(* IEC 61131-3 sources: RVM_Dijital_Ikiz_ModelveOtomasyon_BitirmeProjesi/Codesys_Dosyalari/Paylasim/PLC_Kaynaklari, 10 files *)

(* ---- FB_CikisKontrolLD_decl.st ---- *)
FUNCTION_BLOCK FB_CikisKontrolLD
VAR_INPUT
    // Diagnostic inputs: confirm scan updates without changing ladder logic.
    udiCevrimNo : UDINT;
    uiMakineDurumu : UINT;
	xCalismaIzni: BOOL;
	xBaglanti: BOOL;
	xVeriGecerli: BOOL;
	xAcilStop: BOOL;
	xSikisma: BOOL;
	xDurdur: BOOL;
	xGirisAsamasi: BOOL;
	xKabulAsamasi: BOOL;
	xIadeAsamasi: BOOL;
	xKirmaAsamasi: BOOL;
	xHazneAsamasi: BOOL;
	xEveDonusAsamasi: BOOL;
	xBosaltmaAsamasi: BOOL;
	xTanimaOnayi: BOOL;
	xKapakKapali: BOOL;
	xHedefte: BOOL;
END_VAR
VAR_OUTPUT
	xHareketIzni: BOOL;
	xIleriIstegi: BOOL;
	xGeriIstegi: BOOL;
	xKiriciCalis: BOOL;
	xHazneHareket: BOOL;
	xKapakAc: BOOL;
END_VAR

(* ---- FB_KomutOnceligi106_decl.st ---- *)
FUNCTION_BLOCK FB_KomutOnceligi106
VAR_INPUT
    uiKomutKodu : UINT;
    xYeniKomut : BOOL;
    udiKomutKimligi : UDINT;
END_VAR
VAR_OUTPUT
    uiOncelik : UINT;
    udiCevrimSayaci : UDINT;
    uiSonKomutKodu : UINT;
    uiSonOncelik : UINT;
    udiSonKomutKimligi : UDINT;
END_VAR

(* ---- FB_KonveyorIzin_decl.st ---- *)
FUNCTION_BLOCK FB_KonveyorIzin
VAR_INPUT
    xIzin        : BOOL;
    xIleriIstegi : BOOL;
    xGeriIstegi  : BOOL;
END_VAR
VAR_OUTPUT
    xIleri        : BOOL;
    xGeri         : BOOL;
    xYonCakismasi : BOOL;
END_VAR

(* ---- FB_MalzemeSiniflandirma106_decl.st ---- *)
FUNCTION_BLOCK FB_MalzemeSiniflandirma106
VAR_INPUT
    rMetal : REAL;
    rManyetik : REAL;
    rKutleGram : REAL;
    rGecirgenlik : REAL;
    rYansima : REAL;
    rBoyMetre : REAL;
    rEnMetre : REAL;
    rDoluluk : REAL;
    xVeriYasiUygun : BOOL := TRUE;
    xSensorlerGecerli : BOOL := TRUE;
    xSekilUygun : BOOL := TRUE;
    udiUrunKimligi : UDINT;
    udiPlcOturumu : UDINT;
    udiUnityOturumu : UDINT;
    udiGoruntuIstegi : UDINT;
END_VAR
VAR_OUTPUT
    xDegerlendirildi : BOOL;
    udiDegerlendirmeSayaci : UDINT;
    uiMalzeme : UINT;
    uiGoruntuKarari : UINT;
    uiRetNedeni : UINT;
    rBoyCm : REAL;
    rEnCm : REAL;
    rYuzeyAlani : REAL;
    rHacim : REAL;
    rKabukYogunluk : REAL;
    rHacimYogunluk : REAL;
    xTemelSinirlarUygun : BOOL;
    xAlanUygun : BOOL;
    xPetKosullari : BOOL;
    xCamKosullari : BOOL;
    xAluminyumKosullari : BOOL;
    xMetalBelirsiz : BOOL;
END_VAR

(* ---- FB_RVMControl106_decl.st ---- *)
FUNCTION_BLOCK FB_RVMControl106
VAR_INPUT
    inp : ST_RVMInput106;
    op : ST_RVMOperator106;
    fresh : BOOL;
    epoch : UDINT;
END_VAR
VAR_OUTPUT
    q : ST_RVMOutput106;
END_VAR
VAR
    a : ST_RVMInput106;
    initialized : BOOL;
    session : UDINT;
    packet : UDINT;
    heartbeat : BOOL;
    synchronized : BOOL;
    sessionChanged : BOOL;
    dataOK : BOOL;
    linked : BOOL;
    home : BOOL;
    emptyHome : BOOL;
    emergency : BOOL;
    stopLevel : BOOL;
    targetFull : BOOL;
    faultNow : UINT;
    previousState : UINT;
    previousButtons : ARRAY[1..5] OF BOOL;
    armed : ARRAY[1..5] OF BOOL;
    buttons : ARRAY[1..5] OF BOOL;
    edges : ARRAY[1..5] OF BOOL;
    newRequest : ARRAY[1..2] OF BOOL;
    cmdId : ARRAY[1..2] OF UDINT;
    cmdCode : ARRAY[1..2] OF UINT;
    cmdParam : ARRAY[1..2] OF UINT;
    cachedStatus : ARRAY[1..2] OF UINT;
    cachedReason : ARRAY[1..2] OF UINT;
    replyId : ARRAY[1..2] OF UDINT;
    replyStatus : ARRAY[1..2] OF UINT;
    replyReason : ARRAY[1..2] OF UINT;
    source : INT;
    chosen : INT;
    other : INT;
    i : INT;
    hmiCode : UINT;
    hmiParam : UINT;
    resultStatus : UINT;
    resultReason : UINT;
    pendingSource : INT;
    pendingId : UDINT;
    insertConfirmed : BOOL;
    confirmedProduct : UDINT;
    lastProduct : UDINT;
    waitLink : TON;
    waitStage : TON;
    waitRecognition : TON;
    waitVision : TON;
    visionMatch : BOOL;
    visionShape : BOOL;
    waitCycle : TON;
    waitInsert : TON;
    fbMalzeme : FB_MalzemeSiniflandirma106;
    fbUnityOncelik : FB_KomutOnceligi106;
    fbCodesysOncelik : FB_KomutOnceligi106;
    fbCikisLD : FB_CikisKontrolLD;
    fbKonveyorIzin : FB_KonveyorIzin;
END_VAR

(* ---- FB_KomutOnceligi106_body.st ---- *)
// Same command priorities; separate instances for Unity and CODESYS HMI.
CASE uiKomutKodu OF
2: uiOncelik := 1;
3: uiOncelik := 2;
5: uiOncelik := 3;
1: uiOncelik := 4;
4: uiOncelik := 5;
ELSE uiOncelik := 99;
END_CASE;
IF udiCevrimSayaci = UDINT#4294967295 THEN
    udiCevrimSayaci := 1;
ELSE
    udiCevrimSayaci := udiCevrimSayaci + 1;
END_IF;
IF xYeniKomut THEN
    uiSonKomutKodu := uiKomutKodu;
    uiSonOncelik := uiOncelik;
    udiSonKomutKimligi := udiKomutKimligi;
END_IF;

(* ---- FB_MalzemeSiniflandirma106_body.st ---- *)
// Last completed classification attempt. Inputs and results remain visible.
// Each attempt clears intermediate values, including early rejection paths.
xDegerlendirildi := TRUE;
IF udiDegerlendirmeSayaci = UDINT#4294967295 THEN
    udiDegerlendirmeSayaci := 1;
ELSE
    udiDegerlendirmeSayaci := udiDegerlendirmeSayaci + 1;
END_IF;
uiMalzeme := 0; uiGoruntuKarari := 2; uiRetNedeni := 0;
rBoyCm := 0; rEnCm := 0; rYuzeyAlani := 0; rHacim := 0;
rKabukYogunluk := 0; rHacimYogunluk := 0;
xTemelSinirlarUygun := FALSE; xAlanUygun := FALSE;
xPetKosullari := FALSE; xCamKosullari := FALSE;
xAluminyumKosullari := FALSE; xMetalBelirsiz := FALSE;

// Same order as the previous controller guards.
IF NOT xVeriYasiUygun THEN uiRetNedeni := 10; uiGoruntuKarari := 4; RETURN; END_IF;
IF NOT xSensorlerGecerli THEN uiRetNedeni := 11; uiGoruntuKarari := 3; RETURN; END_IF;
IF NOT xSekilUygun THEN uiRetNedeni := 12; RETURN; END_IF;

xTemelSinirlarUygun := (rMetal>=0) AND (rMetal<=1) AND (rManyetik>=0) AND (rManyetik<=0.1)
    AND (rKutleGram>=5) AND (rKutleGram<=1000) AND (rGecirgenlik>=0) AND (rGecirgenlik<=1)
    AND (rYansima>=0) AND (rYansima<=1) AND (rBoyMetre>=0.10) AND (rBoyMetre<=0.30)
    AND (rEnMetre>=0.02) AND (rEnMetre<=0.09) AND (rDoluluk>0) AND (rDoluluk<=1);
IF NOT xTemelSinirlarUygun THEN uiRetNedeni := 1; RETURN; END_IF;
rBoyCm := rBoyMetre * 100.0;
rEnCm := rEnMetre * 100.0;
rYuzeyAlani := 3.14159265 * rEnCm * rBoyCm * rDoluluk;
xAlanUygun := rYuzeyAlani > 1.0;
IF NOT xAlanUygun THEN uiRetNedeni := 2; RETURN; END_IF;
rHacim := rYuzeyAlani * rEnCm / 4.0;
rKabukYogunluk := rKutleGram / rYuzeyAlani;
rHacimYogunluk := rKutleGram / rHacim;

xAluminyumKosullari := (rMetal>=0.5) AND (rGecirgenlik<=0.08)
    AND (rKutleGram>=8) AND (rKutleGram<=45) AND (rBoyMetre<=0.20);
xPetKosullari := (rMetal<=0.1) AND (rKutleGram>=8) AND (rKutleGram<=75)
    AND (rKabukYogunluk>=0.040) AND (rKabukYogunluk<=0.095) AND (rGecirgenlik>=0.35);
xCamKosullari := (rMetal<=0.1) AND (rKutleGram>=100) AND (rKutleGram<=800)
    AND (rKabukYogunluk>=0.450) AND (rKabukYogunluk<=0.680) AND (rDoluluk>=0.875)
    AND (rGecirgenlik>=0.45) AND (rGecirgenlik<=0.85) AND (rYansima>=0.12);
xMetalBelirsiz := (rMetal>0.1) AND (rMetal<0.5);
IF rMetal>=0.5 THEN
    IF xAluminyumKosullari THEN uiMalzeme := 2; ELSE uiRetNedeni := 3; END_IF;
ELSIF rMetal<=0.1 THEN
    IF xPetKosullari THEN uiMalzeme := 1;
    ELSIF xCamKosullari THEN uiMalzeme := 3;
    ELSE uiRetNedeni := 5;
    END_IF;
ELSE
    uiRetNedeni := 4;
END_IF;
IF uiMalzeme<>0 THEN uiGoruntuKarari := 1; END_IF;

(* ---- FB_RVMControl106_body.st ---- *)
// Single process owner. No actuator command is derived from a UI bit directly.
q.uiProtokolSurumu := 106;
q.udiPlcOturumu := epoch;
q.uiDesteklenenModlar := 2; // Render camera + simulated physical sensors only.
q.uiVeriModu := 1;
q.rBantHizi := 0.85;
q.rKiriciDevri := 120.0;
q.rHazneHizi := 1.5;
q.rKapakAcisi := 75.0;
q.udiPlcSayaci := q.udiPlcSayaci + 1;
heartbeat := FALSE;
sessionChanged := FALSE;
newRequest[1] := FALSE;
newRequest[2] := FALSE;
insertConfirmed := FALSE;
faultNow := 0;
IF NOT initialized THEN
    initialized := TRUE;
    q.uiDurum := 0;
    q.xCalismaIzni := FALSE;
    q.rHazneHedefi := 0.225;
END_IF;
IF epoch = 0 THEN faultNow := 313; END_IF;

// A zero-epoch HELLO is mandatory before this PLC incarnation accepts commands.
// The HELLO'inp command watermark is consumed, never executed.
IF fresh AND (inp.udiUnityOturumu <> 0) AND (inp.udiUnitySayaci <> 0) THEN
    IF (inp.udiGorulenPlcOturumu = 0) AND ((session <> inp.udiUnityOturumu) OR NOT synchronized) THEN
        a := inp;
        sessionChanged := session <> inp.udiUnityOturumu;
        session := inp.udiUnityOturumu;
        lastProduct := 0;
        packet := inp.udiUnitySayaci;
        synchronized := TRUE;
        cmdId[1] := inp.udiKomutKimligi;
        cmdCode[1] := inp.uiOperatorKomutu;
        cmdParam[1] := inp.uiOperatorParametresi;
        cachedStatus[1] := 5;
        cachedReason[1] := 10;
        replyId[1] := cmdId[1];
        replyStatus[1] := 5;
        replyReason[1] := 10;
        q.xCalismaIzni := FALSE;
        IF q.uiHataKodu = 0 THEN q.uiDurum := 0; END_IF;
    ELSIF synchronized AND (session = inp.udiUnityOturumu)
        AND (inp.udiGorulenPlcOturumu = epoch) AND (inp.udiUnitySayaci > packet) THEN
        packet := inp.udiUnitySayaci;
        a := inp;
        heartbeat := TRUE;
        IF inp.udiKomutKimligi > cmdId[1] THEN
            cmdId[1] := inp.udiKomutKimligi;
            cmdCode[1] := inp.uiOperatorKomutu;
            cmdParam[1] := inp.uiOperatorParametresi;
            newRequest[1] := TRUE;
        ELSIF (inp.udiKomutKimligi <> cmdId[1]) OR (inp.uiOperatorKomutu <> cmdCode[1])
            OR (inp.uiOperatorParametresi <> cmdParam[1]) THEN
            replyId[1] := inp.udiKomutKimligi;
            replyStatus[1] := 3;
            replyReason[1] := 13;
        ELSE
            replyId[1] := cmdId[1];
            replyStatus[1] := cachedStatus[1];
            replyReason[1] := cachedReason[1];
        END_IF;
    END_IF;
END_IF;
q.udiUnityOnayOturumu := session;
waitLink(IN := NOT heartbeat, PT := T#750MS);
linked := synchronized AND (session = a.udiUnityOturumu) AND (a.udiGorulenPlcOturumu = epoch)
    AND (epoch <> 0) AND NOT waitLink.Q AND (a.uiUnityProtokol = 106);
home := ABS(a.rHazneKonumu - 0.225) < 0.008;
emptyHome := a.xYolBos AND NOT a.xGiris AND a.xKapakKapali AND NOT a.xKapakAcik AND home;
emergency := op.xAcilStop OR a.xAcilStop;
// Comparisons reject NaN as well as out-of-range values. No invalid data fallback.
dataOK := a.xPlantVerisiGecerli AND (a.uiPlantVeriKaynagi = 1)
    AND (a.rHazneKonumu >= -0.770001) AND (a.rHazneKonumu <= 0.310001)
    AND (a.rKutleGram >= 0.0) AND (a.rKutleGram <= 10000.0)
    AND (a.rBoyMetre >= 0.0) AND (a.rBoyMetre <= 2.000001)
    AND (a.rOptikGecirgenlik >= 0.0) AND (a.rOptikGecirgenlik <= 1.000001)
    AND (a.rGercekBantHizi >= -1.200001) AND (a.rGercekBantHizi <= 1.200001)
    AND (a.rGercekKiriciDevri >= 0.0) AND (a.rGercekKiriciDevri <= 180.0001)
    AND NOT (a.xKapakAcik AND a.xKapakKapali)
    AND NOT (a.xYolBos AND a.xGiris) AND (a.uiBosaltilanKutu <= 3);

// HMI: arm only after FALSE has been observed; held or startup TRUE cannot repeat.
buttons[1] := op.xBaslat; buttons[2] := op.xDurdur; buttons[3] := op.xSifirla;
buttons[4] := op.xNesneEkle; buttons[5] := op.xModUygula;
FOR i := 1 TO 5 DO
    IF NOT buttons[i] THEN armed[i] := TRUE; END_IF;
    edges[i] := armed[i] AND buttons[i] AND NOT previousButtons[i];
    previousButtons[i] := buttons[i];
END_FOR;
hmiCode := 0; hmiParam := 0;
IF edges[2] THEN hmiCode := 2;
ELSIF edges[3] THEN hmiCode := 3;
ELSIF edges[5] THEN hmiCode := 5; hmiParam := op.uiSeciliMod;
ELSIF edges[1] THEN hmiCode := 1;
ELSIF edges[4] THEN hmiCode := 4; hmiParam := op.uiSeciliNesne;
END_IF;
IF hmiCode <> 0 THEN
    IF cmdId[2] = UDINT#4294967295 THEN faultNow := 313;
    ELSE
        cmdId[2] := cmdId[2] + 1;
        cmdCode[2] := hmiCode; cmdParam[2] := hmiParam;
        newRequest[2] := TRUE;
    END_IF;
END_IF;
stopLevel := op.xDurdur OR (newRequest[1] AND (cmdCode[1] = 2));

// Fault priority is stable; reconnecting Unity never clears a latched fault.
IF q.xCalismaIzni THEN
    IF emergency THEN faultNow := 303;
    // Unity also raises its local motion interlock on an identity mismatch.
    // Preserve the specific cause while the session is valid, before generic jam/data flags.
    ELSIF linked AND (q.uiDurum >= 20) AND (q.uiDurum <= 100) AND (a.udiUrunKimligi <> q.udiIslemKimligi) THEN faultNow := 305;
    ELSIF a.xSikisma THEN faultNow := 304;
    ELSIF a.uiUnityProtokol <> 106 THEN faultNow := 302;
    ELSIF NOT linked THEN faultNow := 301;
    ELSIF NOT dataOK THEN faultNow := 310;
    END_IF;
END_IF;
waitStage(IN := (q.uiDurum = previousState) AND (q.uiDurum >= 20) AND (q.uiDurum <= 100), PT := T#8S);
previousState := q.uiDurum;
waitRecognition(IN := q.uiDurum = 30, PT := T#200MS);
waitVision(IN := q.uiDurum = 30, PT := T#4S);
visionMatch := (a.udiGoruntuOnayi = q.udiGoruntuIstegi) AND (q.udiGoruntuIstegi <> 0)
    AND (a.udiGoruntuUrunu = q.udiIslemKimligi) AND (a.udiGoruntuPlcOturumu = epoch)
    AND (a.udiGoruntuUnityOturumu = session);
visionShape := a.xGoruntuNesneVar AND (a.rGoruntuBoy >= 0.10) AND (a.rGoruntuBoy <= 0.30)
    AND (a.rGoruntuEn >= 0.02) AND (a.rGoruntuEn <= 0.09)
    AND (a.rGoruntuBoy >= 1.5*a.rGoruntuEn) AND (a.rGoruntuBoy <= 7.0*a.rGoruntuEn)
    AND (a.rGoruntuDoluluk >= 0.35) AND (a.rGoruntuDoluluk <= 1.0);
waitCycle(IN := (q.uiDurum >= 20) AND (q.uiDurum <= 90), PT := T#5600MS);
waitInsert(IN := q.xNesneIstegiEtkin, PT := T#2S);
IF waitStage.Q AND (faultNow = 0) THEN faultNow := 306; END_IF;
IF faultNow <> 0 AND q.uiHataKodu = 0 THEN q.uiHataKodu := faultNow; END_IF;
IF stopLevel OR emergency OR sessionChanged OR (q.uiHataKodu <> 0) THEN
    q.xCalismaIzni := FALSE;
    IF q.uiHataKodu = 0 THEN q.uiDurum := 0; ELSE q.uiDurum := 900; END_IF;
    IF q.xNesneIstegiEtkin THEN
        cachedStatus[pendingSource] := 5; cachedReason[pendingSource] := 1;
        IF replyId[pendingSource] = pendingId THEN
            replyStatus[pendingSource] := 5; replyReason[pendingSource] := 1;
        END_IF;
    END_IF;
    q.xNesneIstegiEtkin := FALSE;
END_IF;

// Arbitration is deterministic. No deferred queue can start work after a stop.
fbUnityOncelik(uiKomutKodu := cmdCode[1], xYeniKomut := newRequest[1], udiKomutKimligi := cmdId[1]);
fbCodesysOncelik(uiKomutKodu := cmdCode[2], xYeniKomut := newRequest[2], udiKomutKimligi := cmdId[2]);
chosen := 0;
IF newRequest[2] THEN chosen := 2; END_IF;
IF newRequest[1] THEN
    IF chosen = 0 THEN chosen := 1;
    ELSIF fbUnityOncelik.uiOncelik < fbCodesysOncelik.uiOncelik THEN chosen := 1;
    END_IF;
END_IF;
FOR source := 1 TO 2 DO
    IF newRequest[source] THEN
        resultStatus := 3; resultReason := 0;
        replyId[source] := cmdId[source];
        IF (source <> chosen) AND NOT (cmdCode[source] = 2) THEN
            IF stopLevel THEN resultReason := 1; ELSE resultReason := 9; END_IF;
        ELSIF cmdCode[source] = 2 THEN
            q.xCalismaIzni := FALSE;
            IF q.uiHataKodu = 0 THEN q.uiDurum := 0; ELSE q.uiDurum := 900; END_IF;
            resultStatus := 2;
        ELSIF (cmdCode[source] = 0) OR (cmdCode[source] > 5)
            OR ((cmdCode[source] <= 3) AND (cmdParam[source] <> 0))
            OR ((cmdCode[source] = 4) AND (cmdParam[source] > 3))
            OR ((cmdCode[source] = 5) AND (cmdParam[source] > 2)) THEN resultReason := 7;
        ELSIF stopLevel THEN resultReason := 1;
        ELSIF emergency OR a.xSikisma THEN resultReason := 5;
        ELSIF NOT linked OR NOT dataOK THEN resultReason := 2;
        ELSIF q.xNesneIstegiEtkin THEN resultReason := 6;
        ELSE
            CASE cmdCode[source] OF
            1:
                IF q.uiHataKodu <> 0 THEN resultReason := 5;
                ELSIF q.uiDurum <> 0 THEN resultReason := 3;
                ELSIF NOT emptyHome THEN resultReason := 4;
                ELSE q.xCalismaIzni := TRUE; q.uiDurum := 10; resultStatus := 2;
                END_IF;
            3:
                IF q.xCalismaIzni OR ((q.uiDurum <> 0) AND (q.uiDurum <> 900)) THEN resultReason := 3;
                ELSIF NOT emptyHome THEN resultReason := 4;
                ELSIF epoch = 0 THEN resultReason := 10;
                ELSE q.uiHataKodu := 0; q.uiDurum := 0; q.xCalismaIzni := FALSE; resultStatus := 2;
                END_IF;
            4:
                IF q.uiHataKodu <> 0 THEN resultReason := 5;
                ELSIF (q.uiDurum <> 10) OR NOT q.xCalismaIzni THEN resultReason := 3;
                ELSIF NOT emptyHome THEN resultReason := 4;
                ELSIF q.udiNesneIstegi = UDINT#4294967295 THEN resultReason := 10;
                ELSE
                    q.udiNesneIstegi := q.udiNesneIstegi + 1;
                    q.uiNesneProfili := cmdParam[source];
                    q.xNesneIstegiEtkin := TRUE;
                    pendingSource := source; pendingId := cmdId[source];
                    resultStatus := 1;
                END_IF;
            5:
                IF cmdParam[source] <> 1 THEN resultReason := 8;
                ELSIF (q.uiDurum <> 0) OR q.xCalismaIzni THEN resultReason := 3;
                ELSIF NOT emptyHome THEN resultReason := 4;
                ELSE q.uiVeriModu := 1; resultStatus := 2;
                END_IF;
            END_CASE;
        END_IF;
        cachedStatus[source] := resultStatus; cachedReason[source] := resultReason;
        replyStatus[source] := resultStatus; replyReason[source] := resultReason;
        IF source = chosen THEN q.uiSonKomutKaynagi := INT_TO_UINT(source); END_IF;
    END_IF;
END_FOR;

// Product admission is tied to the PLC-issued request, not just a presence bit.
IF q.xNesneIstegiEtkin THEN
    resultStatus := 1; resultReason := 0;
    IF waitInsert.Q THEN
        resultStatus := 4; resultReason := 11;
        q.uiHataKodu := 312; // A delayed physical creation must require explicit recovery.
    ELSIF heartbeat AND (a.udiNesneOnayi = q.udiNesneIstegi) THEN
        IF a.uiNesneSonucu = 2 THEN resultStatus := 3; resultReason := 12;
        ELSIF a.uiNesneSonucu = 1 THEN
            IF (a.udiNesneUrunKimligi <> 0) AND (a.udiNesneUrunKimligi = a.udiUrunKimligi)
                AND (a.udiUrunKimligi > lastProduct) AND a.xGiris AND NOT a.xYolBos THEN
                confirmedProduct := a.udiUrunKimligi;
                lastProduct := a.udiUrunKimligi;
                insertConfirmed := TRUE;
                resultStatus := 2;
            ELSE resultStatus := 3; resultReason := 12; q.uiHataKodu := 312;
            END_IF;
        END_IF;
    END_IF;
    IF resultStatus <> 1 THEN
        q.xNesneIstegiEtkin := FALSE;
        IF cmdId[pendingSource] = pendingId THEN
            cachedStatus[pendingSource] := resultStatus; cachedReason[pendingSource] := resultReason;
        END_IF;
        IF replyId[pendingSource] = pendingId THEN
            replyStatus[pendingSource] := resultStatus; replyReason[pendingSource] := resultReason;
        END_IF;
    END_IF;
END_IF;

targetFull := ((q.uiHedefKutu = 1) AND a.xKutuPetDolu)
    OR ((q.uiHedefKutu = 2) AND a.xKutuAluminyumDolu)
    OR ((q.uiHedefKutu = 3) AND a.xKutuCamDolu);
IF q.xCalismaIzni AND (q.uiDurum >= 40) AND (q.uiDurum <= 70) AND targetFull THEN q.uiHataKodu := 308; END_IF;
IF q.uiHataKodu = 0 AND q.xCalismaIzni THEN
    CASE q.uiDurum OF
    10:
        q.xTanimaOnayi := FALSE; q.uiTaninmisMalzeme := 0; q.uiHedefKutu := 0;
        IF insertConfirmed THEN q.udiIslemKimligi := confirmedProduct; q.uiDurum := 20;
        ELSIF NOT a.xYolBos AND NOT q.xNesneIstegiEtkin THEN q.uiHataKodu := 312;
        END_IF;
    20:
        IF a.xTanima THEN
            IF q.udiGoruntuIstegi = UDINT#4294967295 THEN q.uiHataKodu := 313;
            ELSE q.udiGoruntuIstegi := q.udiGoruntuIstegi+1; q.uiGoruntuKarari := 0; q.uiDurum := 30;
            END_IF;
        END_IF;
    30:
        IF NOT a.xTanima THEN q.uiHataKodu := 307;
        ELSIF waitVision.Q THEN
            q.uiGoruntuKarari := 5; q.uiTaninmisMalzeme := 0; q.uiHedefKutu := 0; q.uiDurum := 100;
        ELSIF waitRecognition.Q AND visionMatch THEN
            q.uiTaninmisMalzeme := 0;
            fbMalzeme(
                rMetal := a.rOlcumMetal, rManyetik := a.rOlcumManyetik,
                rKutleGram := a.rKutleGram, rGecirgenlik := a.rOptikGecirgenlik,
                rYansima := a.rOlcumYansima, rBoyMetre := a.rGoruntuBoy,
                rEnMetre := a.rGoruntuEn, rDoluluk := a.rGoruntuDoluluk,
                xVeriYasiUygun := (a.rGoruntuYasiMs >= 0.0) AND (a.rGoruntuYasiMs <= 2000.0),
                xSensorlerGecerli := a.xGoruntuGecerli AND a.xOlcumTartiGecerli AND a.xOlcumProbGecerli,
                xSekilUygun := visionShape,
                udiUrunKimligi := q.udiIslemKimligi, udiPlcOturumu := epoch,
                udiUnityOturumu := a.udiUnityOturumu, udiGoruntuIstegi := q.udiGoruntuIstegi);
            q.uiTaninmisMalzeme := fbMalzeme.uiMalzeme;
            q.uiGoruntuKarari := fbMalzeme.uiGoruntuKarari;
            q.uiHedefKutu := q.uiTaninmisMalzeme;
            CASE q.uiHedefKutu OF
            1: q.rHazneHedefi := -0.23;
            2: q.rHazneHedefi := -0.77;
            3: q.rHazneHedefi := 0.31;
            END_CASE;
            IF q.uiHedefKutu = 0 THEN q.uiDurum := 100;
            ELSIF ((q.uiHedefKutu=1) AND a.xKutuPetDolu) OR ((q.uiHedefKutu=2) AND a.xKutuAluminyumDolu)
                OR ((q.uiHedefKutu=3) AND a.xKutuCamDolu) THEN q.uiHataKodu := 308;
            ELSE q.xTanimaOnayi := TRUE; q.uiDurum := 40;
            END_IF;
        END_IF;
    40:
        IF NOT a.xKapakKapali THEN q.uiHataKodu := 310;
        ELSIF a.xKiriciGiris THEN q.uiDurum := 50; END_IF;
    50:
        IF a.xKirildi AND a.xHazneDolu AND a.xKapakKapali THEN q.uiDurum := 60; END_IF;
    60:
        IF NOT a.xKapakKapali OR NOT a.xHazneDolu THEN q.uiHataKodu := 310;
        ELSIF ABS(a.rHazneKonumu-q.rHazneHedefi)<0.008 THEN q.uiDurum := 70; END_IF;
    70:
        IF ABS(a.rHazneKonumu-q.rHazneHedefi)>=0.008 THEN q.uiHataKodu := 310;
        ELSIF a.xBosaltildi AND a.xKapakAcik AND NOT a.xHazneDolu AND a.xYolBos THEN
            IF a.uiBosaltilanKutu <> q.uiHedefKutu THEN q.uiHataKodu := 309;
            ELSE q.uiDurum := 80; END_IF;
        END_IF;
    80:
        IF a.xKapakKapali AND NOT a.xKapakAcik AND a.xYolBos AND NOT a.xHazneDolu THEN
            CASE q.uiHedefKutu OF
            1: q.udiPetSayaci := q.udiPetSayaci + 1;
            2: q.udiAluminyumSayaci := q.udiAluminyumSayaci + 1;
            3: q.udiCamSayaci := q.udiCamSayaci + 1;
            END_CASE;
            q.uiDurum := 90;
        END_IF;
    90:
        q.rHazneHedefi := 0.225;
        IF NOT a.xKapakKapali THEN q.uiHataKodu := 310;
        ELSIF home AND a.xYolBos AND waitCycle.Q THEN q.uiDurum := 10; END_IF;
    100:
        IF a.xYolBos THEN q.udiReddedilenSayaci := q.udiReddedilenSayaci+1; q.uiDurum := 10; END_IF;
    END_CASE;
END_IF;

// Apply fault dominance AFTER state processing, in this same scan.
IF q.uiHataKodu <> 0 THEN q.uiDurum := 900; q.xCalismaIzni := FALSE; q.xNesneIstegiEtkin := FALSE; END_IF;
fbCikisLD(
    udiCevrimNo := q.udiPlcSayaci, uiMakineDurumu := q.uiDurum,
    xCalismaIzni := q.xCalismaIzni, xBaglanti := linked, xVeriGecerli := dataOK,
    xAcilStop := emergency, xSikisma := a.xSikisma, xDurdur := stopLevel,
    xGirisAsamasi := q.uiDurum=20, xKabulAsamasi := q.uiDurum=40,
    xIadeAsamasi := q.uiDurum=100, xKirmaAsamasi := q.uiDurum=50,
    xHazneAsamasi := q.uiDurum=60, xEveDonusAsamasi := q.uiDurum=90,
    xBosaltmaAsamasi := q.uiDurum=70, xTanimaOnayi := q.xTanimaOnayi,
    xKapakKapali := a.xKapakKapali, xHedefte := ABS(a.rHazneKonumu-q.rHazneHedefi)<0.008);
fbKonveyorIzin(xIzin := fbCikisLD.xHareketIzni,
    xIleriIstegi := fbCikisLD.xIleriIstegi, xGeriIstegi := fbCikisLD.xGeriIstegi);
q.xKonveyorIleri := fbKonveyorIzin.xIleri;
q.xKonveyorGeri := fbKonveyorIzin.xGeri;
q.xKiriciCalis := fbCikisLD.xKiriciCalis;
q.xHazneHareket := fbCikisLD.xHazneHareket;
q.xKapakAc := fbCikisLD.xKapakAc;
IF NOT q.xCalismaIzni THEN q.xTanimaOnayi := FALSE; END_IF;
q.udiKomutOnayi := replyId[1]; q.uiKomutDurumu := replyStatus[1]; q.uiKomutNedeni := replyReason[1];
q.udiPlcOperatorKomutKimligi := replyId[2]; q.uiPlcOperatorKomutu := cmdCode[2];
q.uiPlcKomutDurumu := replyStatus[2]; q.uiPlcKomutNedeni := replyReason[2];

(* ---- PRG_UnityRVM_body.st ---- *)
IF NOT initialized THEN
    initialized := TRUE;
    IF GVL_RVMKalici.udiOturum < UDINT#4294967295 THEN
        GVL_RVMKalici.udiOturum := GVL_RVMKalici.udiOturum + 1;
        epoch := GVL_RVMKalici.udiOturum;
    END_IF;
END_IF;
fresh := FALSE;
beginMarker := GVL_RVMUnity.udiGirisBaslangic;
IF (beginMarker <> 0) AND (beginMarker = GVL_RVMUnity.udiGirisBitis) AND (beginMarker <> lastMarker) THEN
candidate.uiUnityProtokol := GVL_RVMUnity.uiUnityProtokol;
candidate.udiUnityOturumu := GVL_RVMUnity.udiUnityOturumu;
candidate.udiUnitySayaci := GVL_RVMUnity.udiUnitySayaci;
candidate.udiKomutKimligi := GVL_RVMUnity.udiKomutKimligi;
candidate.uiOperatorKomutu := GVL_RVMUnity.uiOperatorKomutu;
candidate.xGiris := GVL_RVMUnity.xGiris;
candidate.xTanima := GVL_RVMUnity.xTanima;
candidate.xKiriciGiris := GVL_RVMUnity.xKiriciGiris;
candidate.xKirildi := GVL_RVMUnity.xKirildi;
candidate.xHazneDolu := GVL_RVMUnity.xHazneDolu;
candidate.xBosaltildi := GVL_RVMUnity.xBosaltildi;
candidate.xKapakAcik := GVL_RVMUnity.xKapakAcik;
candidate.xKapakKapali := GVL_RVMUnity.xKapakKapali;
candidate.xYolBos := GVL_RVMUnity.xYolBos;
candidate.xMetalAlgilandi := GVL_RVMUnity.xMetalAlgilandi;
candidate.xSikisma := GVL_RVMUnity.xSikisma;
candidate.xAcilStop := GVL_RVMUnity.xAcilStop;
candidate.xKutuPetDolu := GVL_RVMUnity.xKutuPetDolu;
candidate.xKutuAluminyumDolu := GVL_RVMUnity.xKutuAluminyumDolu;
candidate.xKutuCamDolu := GVL_RVMUnity.xKutuCamDolu;
candidate.rKutleGram := GVL_RVMUnity.rKutleGram;
candidate.rOptikGecirgenlik := GVL_RVMUnity.rOptikGecirgenlik;
candidate.rBoyMetre := GVL_RVMUnity.rBoyMetre;
candidate.rHazneKonumu := GVL_RVMUnity.rHazneKonumu;
candidate.rGercekBantHizi := GVL_RVMUnity.rGercekBantHizi;
candidate.rGercekKiriciDevri := GVL_RVMUnity.rGercekKiriciDevri;
candidate.uiBosaltilanKutu := GVL_RVMUnity.uiBosaltilanKutu;
candidate.udiUrunKimligi := GVL_RVMUnity.udiUrunKimligi;
candidate.uiOperatorParametresi := GVL_RVMUnity.uiOperatorParametresi;
candidate.udiGorulenPlcOturumu := GVL_RVMUnity.udiGorulenPlcOturumu;
candidate.udiNesneOnayi := GVL_RVMUnity.udiNesneOnayi;
candidate.uiNesneSonucu := GVL_RVMUnity.uiNesneSonucu;
candidate.udiNesneUrunKimligi := GVL_RVMUnity.udiNesneUrunKimligi;
candidate.uiPlantVeriKaynagi := GVL_RVMUnity.uiPlantVeriKaynagi;
candidate.xPlantVerisiGecerli := GVL_RVMUnity.xPlantVerisiGecerli;
candidate.udiGoruntuOnayi := GVL_RVMUnity.udiGoruntuOnayi;
candidate.udiGoruntuUrunu := GVL_RVMUnity.udiGoruntuUrunu;
candidate.udiGoruntuPlcOturumu := GVL_RVMUnity.udiGoruntuPlcOturumu;
candidate.udiGoruntuUnityOturumu := GVL_RVMUnity.udiGoruntuUnityOturumu;
candidate.xGoruntuGecerli := GVL_RVMUnity.xGoruntuGecerli;
candidate.xGoruntuNesneVar := GVL_RVMUnity.xGoruntuNesneVar;
candidate.rGoruntuBoy := GVL_RVMUnity.rGoruntuBoy;
candidate.rGoruntuEn := GVL_RVMUnity.rGoruntuEn;
candidate.rGoruntuDoluluk := GVL_RVMUnity.rGoruntuDoluluk;
candidate.rGoruntuYasiMs := GVL_RVMUnity.rGoruntuYasiMs;
candidate.xOlcumTartiGecerli := GVL_RVMUnity.xOlcumTartiGecerli;
candidate.xOlcumProbGecerli := GVL_RVMUnity.xOlcumProbGecerli;
candidate.rOlcumYansima := GVL_RVMUnity.rOlcumYansima;
candidate.rOlcumMetal := GVL_RVMUnity.rOlcumMetal;
candidate.rOlcumManyetik := GVL_RVMUnity.rOlcumManyetik;
    fresh := (beginMarker = GVL_RVMUnity.udiGirisBitis) AND (beginMarker = GVL_RVMUnity.udiGirisBaslangic);
    IF fresh THEN snapshot := candidate; lastMarker := beginMarker; END_IF;
END_IF;
op.xBaslat := GVL_RVMOperator.xBaslat;
op.xDurdur := GVL_RVMOperator.xDurdur;
op.xSifirla := GVL_RVMOperator.xSifirla;
op.xNesneEkle := GVL_RVMOperator.xNesneEkle;
op.xModUygula := GVL_RVMOperator.xModUygula;
op.xAcilStop := GVL_RVMOperator.xAcilStop;
op.uiSeciliNesne := GVL_RVMOperator.uiSeciliNesne;
op.uiSeciliMod := GVL_RVMOperator.uiSeciliMod;
control(inp := snapshot, op := op, fresh := fresh, epoch := epoch);
IF outputMarker = UDINT#4294967295 THEN outputMarker := 1; ELSE outputMarker := outputMarker+1; END_IF;
GVL_RVMUnity.udiCikisBaslangic := outputMarker;
GVL_RVMUnity.uiProtokolSurumu := control.q.uiProtokolSurumu;
GVL_RVMUnity.udiPlcSayaci := control.q.udiPlcSayaci;
GVL_RVMUnity.udiUnityOnayOturumu := control.q.udiUnityOnayOturumu;
GVL_RVMUnity.udiGirisOnayi := control.q.udiGirisOnayi;
GVL_RVMUnity.udiKomutOnayi := control.q.udiKomutOnayi;
GVL_RVMUnity.udiIslemKimligi := control.q.udiIslemKimligi;
GVL_RVMUnity.uiDurum := control.q.uiDurum;
GVL_RVMUnity.uiHataKodu := control.q.uiHataKodu;
GVL_RVMUnity.uiTaninmisMalzeme := control.q.uiTaninmisMalzeme;
GVL_RVMUnity.uiHedefKutu := control.q.uiHedefKutu;
GVL_RVMUnity.xCalismaIzni := control.q.xCalismaIzni;
GVL_RVMUnity.xKonveyorIleri := control.q.xKonveyorIleri;
GVL_RVMUnity.xKonveyorGeri := control.q.xKonveyorGeri;
GVL_RVMUnity.xKiriciCalis := control.q.xKiriciCalis;
GVL_RVMUnity.xHazneHareket := control.q.xHazneHareket;
GVL_RVMUnity.xKapakAc := control.q.xKapakAc;
GVL_RVMUnity.xTanimaOnayi := control.q.xTanimaOnayi;
GVL_RVMUnity.rBantHizi := control.q.rBantHizi;
GVL_RVMUnity.rKiriciDevri := control.q.rKiriciDevri;
GVL_RVMUnity.rHazneHizi := control.q.rHazneHizi;
GVL_RVMUnity.rHazneHedefi := control.q.rHazneHedefi;
GVL_RVMUnity.rKapakAcisi := control.q.rKapakAcisi;
GVL_RVMUnity.udiPetSayaci := control.q.udiPetSayaci;
GVL_RVMUnity.udiAluminyumSayaci := control.q.udiAluminyumSayaci;
GVL_RVMUnity.udiCamSayaci := control.q.udiCamSayaci;
GVL_RVMUnity.udiReddedilenSayaci := control.q.udiReddedilenSayaci;
GVL_RVMUnity.udiPlcOturumu := control.q.udiPlcOturumu;
GVL_RVMUnity.uiKomutDurumu := control.q.uiKomutDurumu;
GVL_RVMUnity.uiKomutNedeni := control.q.uiKomutNedeni;
GVL_RVMUnity.udiPlcOperatorKomutKimligi := control.q.udiPlcOperatorKomutKimligi;
GVL_RVMUnity.uiPlcOperatorKomutu := control.q.uiPlcOperatorKomutu;
GVL_RVMUnity.uiPlcKomutDurumu := control.q.uiPlcKomutDurumu;
GVL_RVMUnity.uiPlcKomutNedeni := control.q.uiPlcKomutNedeni;
GVL_RVMUnity.uiSonKomutKaynagi := control.q.uiSonKomutKaynagi;
GVL_RVMUnity.udiNesneIstegi := control.q.udiNesneIstegi;
GVL_RVMUnity.uiNesneProfili := control.q.uiNesneProfili;
GVL_RVMUnity.xNesneIstegiEtkin := control.q.xNesneIstegiEtkin;
GVL_RVMUnity.uiVeriModu := control.q.uiVeriModu;
GVL_RVMUnity.uiDesteklenenModlar := control.q.uiDesteklenenModlar;
GVL_RVMUnity.udiGoruntuIstegi := control.q.udiGoruntuIstegi;
GVL_RVMUnity.uiGoruntuKarari := control.q.uiGoruntuKarari;
GVL_RVMUnity.udiGirisOnayi := lastMarker;
GVL_RVMUnity.udiCikisBitis := outputMarker;

(* ---- PRG_UnityRVM_decl.st ---- *)
PROGRAM PRG_UnityRVM
VAR
    control : FB_RVMControl106;
    candidate : ST_RVMInput106;
    snapshot : ST_RVMInput106;
    op : ST_RVMOperator106;
    initialized : BOOL;
    epoch : UDINT;
    beginMarker : UDINT;
    lastMarker : UDINT;
    outputMarker : UDINT;
    fresh : BOOL;
END_VAR
